Fanuc KAREL source: kf00054.KL

-- PROVISIONAL review KL for V940-1; original PC SHA256 192c4a62282f60f694cbe043900961266722d3f1b28679d50cb0c29fe955e287
-- Incomplete behavior may be omitted. Consult companion uncertainty JSON. Do not deploy.
PROGRAM KF00054
%NOLOCKGROUP
VAR
  I : INTEGER
  J : INTEGER
  X : REAL
  Y : REAL
  B : BOOLEAN
  C : BOOLEAN
  TXT : STRING[80]
  TXT2 : STRING[80]
  STATUS : INTEGER
-- UNRESOLVED_DECL AI type=002010
-- UNRESOLVED_DECL BI type=002010
-- UNRESOLVED_DECL P type=000102
-- UNRESOLVED_DECL JP type=000199
-- UNRESOLVED_DECL PF type=000101
-- UNRESOLVED_DECL V1 type=000013
-- UNRESOLVED_DECL V2 type=000013
BEGIN
  -- V9_EXPOSED_INDEXED_TABLE_HINT layout=0001; 1 counted words exposed once; source arms/runtime held
  -- UNRESOLVED_PC offsets 5-12; opcodes 9D,23
  -- UNRESOLVED_PC offsets 17-22; opcodes 7A
  -- UNRESOLVED_PC offsets 27-38; opcodes 2E,23
  -- UNRESOLVED_PC offsets 43-54; opcodes 2E,23
  -- UNRESOLVED_PC offsets 59-63; opcodes 7F
END KF00054
